Fanuc KAREL source: compact_preamble.KL

PROGRAM KA00027
%NOLOCKGROUP
VAR
SRC:BOOLEAN;DST:BOOLEAN
BEGIN
SRC=TRUE
DST=SRC
END KA00027
